(* IEC 61131-3 sources: plc-st-coding-agent/progress/evidence/f14_v5_public_pilot_20261112/jobs/custom_deepseek-v4pro, 22 files *)

(* ---- public-easy-01.candidate_01.st ---- *)
TYPE LineState :
(
    IDLE,
    CLEANING,
    FILLING,
    CAPPING,
    PACKING,
    COMPLETE
);
END_TYPE;

FUNCTION_BLOCK AutomatedFillingLine
VAR_INPUT
    bottleSensor : BOOL;
    cleaningConfirmButton : BOOL;
    fillingConfirmButton : BOOL;
    cappingConfirmButton : BOOL;
    packingConfirmButton : BOOL;
    finishedButton : BOOL;
END_VAR
VAR_OUTPUT
    Pump_Motor : BOOL;
    Filling_Valve : BOOL;
    Capping_Machine : BOOL;
    Packing_Machine : BOOL;
    Completion_Light : BOOL;
END_VAR
VAR
    cleaningEdge : R_TRIG;
    fillingEdge : R_TRIG;
    cappingEdge : R_TRIG;
    packingEdge : R_TRIG;
    finishedEdge : R_TRIG;
    currentState : LineState := LineState#IDLE;
END_VAR

(*
ENGINEERING_CONTRACT
- Pump_Motor: activated when bottleSensor TRUE and state=IDLE -> CLEANING; retained until cleaningConfirm edge (PUB003, PUB004).
  Deactivated on cleaningConfirm edge.
- Filling_Valve: activated on cleaningConfirm edge after cleaning; retained until fillingConfirm edge (PUB004, PUB005).
  Deactivated on fillingConfirm edge.
- Capping_Machine: activated on fillingConfirm edge; retained until cappingConfirm edge (PUB005, PUB006).
  Deactivated on cappingConfirm edge.
- Packing_Machine: activated on cappingConfirm edge; retained until packingConfirm edge (PUB006, PUB007).
  Deactivated on packingConfirm edge.
- Completion_Light: activated on packingConfirm edge; retained until finishedButton edge (PUB007, PUB008).
  Deactivated on finishedButton edge, which also resets state to IDLE for next bottle.
- Same-scan priority: state transitions evaluated sequentially in scan order; no simultaneous edge trigger priority specified.
- Units: BOOL levels only; no timing/modbus scaling.
*)

cleaningEdge(CLK := cleaningConfirmButton);
fillingEdge(CLK := fillingConfirmButton);
cappingEdge(CLK := cappingConfirmButton);
packingEdge(CLK := packingConfirmButton);
finishedEdge(CLK := finishedButton);

CASE currentState OF
    LineState#IDLE:
        Pump_Motor := FALSE;
        Filling_Valve := FALSE;
        Capping_Machine := FALSE;
        Packing_Machine := FALSE;
        Completion_Light := FALSE;

        IF bottleSensor THEN
            currentState := LineState#CLEANING;
            Pump_Motor := TRUE;
        END_IF;

    LineState#CLEANING:
        Pump_Motor := TRUE;
        Filling_Valve := FALSE;
        Capping_Machine := FALSE;
        Packing_Machine := FALSE;
        Completion_Light := FALSE;

        IF cleaningEdge.Q THEN
            Pump_Motor := FALSE;
            Filling_Valve := TRUE;
            currentState := LineState#FILLING;
        END_IF;

    LineState#FILLING:
        Pump_Motor := FALSE;
        Filling_Valve := TRUE;
        Capping_Machine := FALSE;
        Packing_Machine := FALSE;
        Completion_Light := FALSE;

        IF fillingEdge.Q THEN
            Filling_Valve := FALSE;
            Capping_Machine := TRUE;
            currentState := LineState#CAPPING;
        END_IF;

    LineState#CAPPING:
        Pump_Motor := FALSE;
        Filling_Valve := FALSE;
        Capping_Machine := TRUE;
        Packing_Machine := FALSE;
        Completion_Light := FALSE;

        IF cappingEdge.Q THEN
            Capping_Machine := FALSE;
            Packing_Machine := TRUE;
            currentState := LineState#PACKING;
        END_IF;

    LineState#PACKING:
        Pump_Motor := FALSE;
        Filling_Valve := FALSE;
        Capping_Machine := FALSE;
        Packing_Machine := TRUE;
        Completion_Light := FALSE;

        IF packingEdge.Q THEN
            Packing_Machine := FALSE;
            Completion_Light := TRUE;
            currentState := LineState#COMPLETE;
        END_IF;

    LineState#COMPLETE:
        Pump_Motor := FALSE;
        Filling_Valve := FALSE;
        Capping_Machine := FALSE;
        Packing_Machine := FALSE;
        Completion_Light := TRUE;

        IF finishedEdge.Q THEN
            Completion_Light := FALSE;
            currentState := LineState#IDLE;
        END_IF;
END_CASE;
END_FUNCTION_BLOCK

(* ---- public-easy-01.candidate_02.st ---- *)
(*
ENGINEERING_CONTRACT
- Pump_Motor: activated when bottleSensor TRUE and state=IDLE -> CLEANING; retained until cleaningConfirm edge (PUB003, PUB004).
  Deactivated on cleaningConfirm edge.
- Filling_Valve: activated on cleaningConfirm edge after cleaning; retained until fillingConfirm edge (PUB004, PUB005).
  Deactivated on fillingConfirm edge.
- Capping_Machine: activated on fillingConfirm edge; retained until cappingConfirm edge (PUB005, PUB006).
  Deactivated on cappingConfirm edge.
- Packing_Machine: activated on cappingConfirm edge; retained until packingConfirm edge (PUB006, PUB007).
  Deactivated on packingConfirm edge.
- Completion_Light: activated on packingConfirm edge; retained until finishedButton edge (PUB007, PUB008).
  Deactivated on finishedButton edge, which also resets state to IDLE for next bottle.
- Same-scan priority: no simultaneous edge trigger priority specified; transitions evaluated sequentially.
- Units: BOOL levels only.
*)

TYPE LineState :
(
    IDLE,
    CLEANING,
    FILLING,
    CAPPING,
    PACKING,
    COMPLETE
);
END_TYPE;

FUNCTION_BLOCK AutomatedFillingLine
VAR_INPUT
    bottleSensor : BOOL;
    cleaningConfirmButton : BOOL;
    fillingConfirmButton : BOOL;
    cappingConfirmButton : BOOL;
    packingConfirmButton : BOOL;
    finishedButton : BOOL;
END_VAR
VAR_OUTPUT
    Pump_Motor : BOOL;
    Filling_Valve : BOOL;
    Capping_Machine : BOOL;
    Packing_Machine : BOOL;
    Completion_Light : BOOL;
END_VAR
VAR
    cleaningEdge : R_TRIG;
    fillingEdge : R_TRIG;
    cappingEdge : R_TRIG;
    packingEdge : R_TRIG;
    finishedEdge : R_TRIG;
    currentState : LineState := IDLE;
END_VAR

cleaningEdge(CLK := cleaningConfirmButton);
fillingEdge(CLK := fillingConfirmButton);
cappingEdge(CLK := cappingConfirmButton);
packingEdge(CLK := packingConfirmButton);
finishedEdge(CLK := finishedButton);

CASE currentState OF
    IDLE:
        Pump_Motor := FALSE;
        Filling_Valve := FALSE;
        Capping_Machine := FALSE;
        Packing_Machine := FALSE;
        Completion_Light := FALSE;

        IF bottleSensor THEN
            currentState := CLEANING;
            Pump_Motor := TRUE;
        END_IF;

    CLEANING:
        Pump_Motor := TRUE;
        Filling_Valve := FALSE;
        Capping_Machine := FALSE;
        Packing_Machine := FALSE;
        Completion_Light := FALSE;

        IF cleaningEdge.Q THEN
            Pump_Motor := FALSE;
            Filling_Valve := TRUE;
            currentState := FILLING;
        END_IF;

    FILLING:
        Pump_Motor := FALSE;
        Filling_Valve := TRUE;
        Capping_Machine := FALSE;
        Packing_Machine := FALSE;
        Completion_Light := FALSE;

        IF fillingEdge.Q THEN
            Filling_Valve := FALSE;
            Capping_Machine := TRUE;
            currentState := CAPPING;
        END_IF;

    CAPPING:
        Pump_Motor := FALSE;
        Filling_Valve := FALSE;
        Capping_Machine := TRUE;
        Packing_Machine := FALSE;
        Completion_Light := FALSE;

        IF cappingEdge.Q THEN
            Capping_Machine := FALSE;
            Packing_Machine := TRUE;
            currentState := PACKING;
        END_IF;

    PACKING:
        Pump_Motor := FALSE;
        Filling_Valve := FALSE;
        Capping_Machine := FALSE;
        Packing_Machine := TRUE;
        Completion_Light := FALSE;

        IF packingEdge.Q THEN
            Packing_Machine := FALSE;
            Completion_Light := TRUE;
            currentState := COMPLETE;
        END_IF;

    COMPLETE:
        Pump_Motor := FALSE;
        Filling_Valve := FALSE;
        Capping_Machine := FALSE;
        Packing_Machine := FALSE;
        Completion_Light := TRUE;

        IF finishedEdge.Q THEN
            Completion_Light := FALSE;
            currentState := IDLE;
        END_IF;
END_CASE;

END_FUNCTION_BLOCK

(* ---- public-easy-01.raw_candidate_01.st ---- *)
TYPE LineState :
(
    IDLE,
    CLEANING,
    FILLING,
    CAPPING,
    PACKING,
    COMPLETE
);
END_TYPE

FUNCTION_BLOCK AutomatedFillingLine
VAR_INPUT
    bottleSensor : BOOL;
    cleaningConfirmButton : BOOL;
    fillingConfirmButton : BOOL;
    cappingConfirmButton : BOOL;
    packingConfirmButton : BOOL;
    finishedButton : BOOL;
END_VAR
VAR_OUTPUT
    Pump_Motor : BOOL;
    Filling_Valve : BOOL;
    Capping_Machine : BOOL;
    Packing_Machine : BOOL;
    Completion_Light : BOOL;
END_VAR
VAR
    cleaningEdge : R_TRIG;
    fillingEdge : R_TRIG;
    cappingEdge : R_TRIG;
    packingEdge : R_TRIG;
    finishedEdge : R_TRIG;
    currentState : LineState := LineState#IDLE;
END_VAR

(*
ENGINEERING_CONTRACT
- Pump_Motor: activated when bottleSensor TRUE and state=IDLE -> CLEANING; retained until cleaningConfirm edge (PUB003, PUB004).
  Deactivated on cleaningConfirm edge.
- Filling_Valve: activated on cleaningConfirm edge after cleaning; retained until fillingConfirm edge (PUB004, PUB005).
  Deactivated on fillingConfirm edge.
- Capping_Machine: activated on fillingConfirm edge; retained until cappingConfirm edge (PUB005, PUB006).
  Deactivated on cappingConfirm edge.
- Packing_Machine: activated on cappingConfirm edge; retained until packingConfirm edge (PUB006, PUB007).
  Deactivated on packingConfirm edge.
- Completion_Light: activated on packingConfirm edge; retained until finishedButton edge (PUB007, PUB008).
  Deactivated on finishedButton edge, which also resets state to IDLE for next bottle.
- Same-scan priority: state transitions evaluated sequentially in scan order; no simultaneous edge trigger priority specified.
- Units: BOOL levels only; no timing/modbus scaling.
*)

cleaningEdge(CLK := cleaningConfirmButton);
fillingEdge(CLK := fillingConfirmButton);
cappingEdge(CLK := cappingConfirmButton);
packingEdge(CLK := packingConfirmButton);
finishedEdge(CLK := finishedButton);

CASE currentState OF
    LineState#IDLE:
        Pump_Motor := FALSE;
        Filling_Valve := FALSE;
        Capping_Machine := FALSE;
        Packing_Machine := FALSE;
        Completion_Light := FALSE;

        IF bottleSensor THEN
            currentState := LineState#CLEANING;
            Pump_Motor := TRUE;
        END_IF;

    LineState#CLEANING:
        Pump_Motor := TRUE;
        Filling_Valve := FALSE;
        Capping_Machine := FALSE;
        Packing_Machine := FALSE;
        Completion_Light := FALSE;

        IF cleaningEdge.Q THEN
            Pump_Motor := FALSE;
            Filling_Valve := TRUE;
            currentState := LineState#FILLING;
        END_IF;

    LineState#FILLING:
        Pump_Motor := FALSE;
        Filling_Valve := TRUE;
        Capping_Machine := FALSE;
        Packing_Machine := FALSE;
        Completion_Light := FALSE;

        IF fillingEdge.Q THEN
            Filling_Valve := FALSE;
            Capping_Machine := TRUE;
            currentState := LineState#CAPPING;
        END_IF;

    LineState#CAPPING:
        Pump_Motor := FALSE;
        Filling_Valve := FALSE;
        Capping_Machine := TRUE;
        Packing_Machine := FALSE;
        Completion_Light := FALSE;

        IF cappingEdge.Q THEN
            Capping_Machine := FALSE;
            Packing_Machine := TRUE;
            currentState := LineState#PACKING;
        END_IF;

    LineState#PACKING:
        Pump_Motor := FALSE;
        Filling_Valve := FALSE;
        Capping_Machine := FALSE;
        Packing_Machine := TRUE;
        Completion_Light := FALSE;

        IF packingEdge.Q THEN
            Packing_Machine := FALSE;
            Completion_Light := TRUE;
            currentState := LineState#COMPLETE;
        END_IF;

    LineState#COMPLETE:
        Pump_Motor := FALSE;
        Filling_Valve := FALSE;
        Capping_Machine := FALSE;
        Packing_Machine := FALSE;
        Completion_Light := TRUE;

        IF finishedEdge.Q THEN
            Completion_Light := FALSE;
            currentState := LineState#IDLE;
        END_IF;
END_CASE;
END_FUNCTION_BLOCK

(* ---- public-easy-01.raw_candidate_02.st ---- *)
(*
ENGINEERING_CONTRACT
- Pump_Motor: activated when bottleSensor TRUE and state=IDLE -> CLEANING; retained until cleaningConfirm edge (PUB003, PUB004).
  Deactivated on cleaningConfirm edge.
- Filling_Valve: activated on cleaningConfirm edge after cleaning; retained until fillingConfirm edge (PUB004, PUB005).
  Deactivated on fillingConfirm edge.
- Capping_Machine: activated on fillingConfirm edge; retained until cappingConfirm edge (PUB005, PUB006).
  Deactivated on cappingConfirm edge.
- Packing_Machine: activated on cappingConfirm edge; retained until packingConfirm edge (PUB006, PUB007).
  Deactivated on packingConfirm edge.
- Completion_Light: activated on packingConfirm edge; retained until finishedButton edge (PUB007, PUB008).
  Deactivated on finishedButton edge, which also resets state to IDLE for next bottle.
- Same-scan priority: no simultaneous edge trigger priority specified; transitions evaluated sequentially.
- Units: BOOL levels only.
*)

TYPE LineState :
(
    IDLE,
    CLEANING,
    FILLING,
    CAPPING,
    PACKING,
    COMPLETE
);
END_TYPE

FUNCTION_BLOCK AutomatedFillingLine
VAR_INPUT
    bottleSensor : BOOL;
    cleaningConfirmButton : BOOL;
    fillingConfirmButton : BOOL;
    cappingConfirmButton : BOOL;
    packingConfirmButton : BOOL;
    finishedButton : BOOL;
END_VAR
VAR_OUTPUT
    Pump_Motor : BOOL;
    Filling_Valve : BOOL;
    Capping_Machine : BOOL;
    Packing_Machine : BOOL;
    Completion_Light : BOOL;
END_VAR
VAR
    cleaningEdge : R_TRIG;
    fillingEdge : R_TRIG;
    cappingEdge : R_TRIG;
    packingEdge : R_TRIG;
    finishedEdge : R_TRIG;
    currentState : LineState := IDLE;
END_VAR

cleaningEdge(CLK := cleaningConfirmButton);
fillingEdge(CLK := fillingConfirmButton);
cappingEdge(CLK := cappingConfirmButton);
packingEdge(CLK := packingConfirmButton);
finishedEdge(CLK := finishedButton);

CASE currentState OF
    IDLE:
        Pump_Motor := FALSE;
        Filling_Valve := FALSE;
        Capping_Machine := FALSE;
        Packing_Machine := FALSE;
        Completion_Light := FALSE;

        IF bottleSensor THEN
            currentState := CLEANING;
            Pump_Motor := TRUE;
        END_IF;

    CLEANING:
        Pump_Motor := TRUE;
        Filling_Valve := FALSE;
        Capping_Machine := FALSE;
        Packing_Machine := FALSE;
        Completion_Light := FALSE;

        IF cleaningEdge.Q THEN
            Pump_Motor := FALSE;
            Filling_Valve := TRUE;
            currentState := FILLING;
        END_IF;

    FILLING:
        Pump_Motor := FALSE;
        Filling_Valve := TRUE;
        Capping_Machine := FALSE;
        Packing_Machine := FALSE;
        Completion_Light := FALSE;

        IF fillingEdge.Q THEN
            Filling_Valve := FALSE;
            Capping_Machine := TRUE;
            currentState := CAPPING;
        END_IF;

    CAPPING:
        Pump_Motor := FALSE;
        Filling_Valve := FALSE;
        Capping_Machine := TRUE;
        Packing_Machine := FALSE;
        Completion_Light := FALSE;

        IF cappingEdge.Q THEN
            Capping_Machine := FALSE;
            Packing_Machine := TRUE;
            currentState := PACKING;
        END_IF;

    PACKING:
        Pump_Motor := FALSE;
        Filling_Valve := FALSE;
        Capping_Machine := FALSE;
        Packing_Machine := TRUE;
        Completion_Light := FALSE;

        IF packingEdge.Q THEN
            Packing_Machine := FALSE;
            Completion_Light := TRUE;
            currentState := COMPLETE;
        END_IF;

    COMPLETE:
        Pump_Motor := FALSE;
        Filling_Valve := FALSE;
        Capping_Machine := FALSE;
        Packing_Machine := FALSE;
        Completion_Light := TRUE;

        IF finishedEdge.Q THEN
            Completion_Light := FALSE;
            currentState := IDLE;
        END_IF;
END_CASE;

END_FUNCTION_BLOCK

(* ---- public-easy-04.candidate_01.st ---- *)
FUNCTION_BLOCK FB_JamPumpDebounceRuntime
VAR_INPUT
    VISCOSITY_OK : BOOL;
    PASTE_E_STOP_NC : BOOL;
    DebounceTime : TIME;
    CycleTime : TIME;
END_VAR
VAR_OUTPUT
    VFD_RUN : BOOL := FALSE;
    PUMP_MAINT_DUE : BOOL := FALSE;
    PUMP_RUNTIME_ACC : LTIME := LTIME#0s;
END_VAR
VAR
    DebounceTimer : TON;
    TonIn : BOOL;
    ViscosityValid : BOOL;
    AccRuntime : LTIME := LTIME#0s;
    MAINT_THRESHOLD : LTIME := LTIME#500h;
END_VAR

(*
ENGINEERING_CONTRACT:
- VFD_RUN activation: PASTE_E_STOP_NC AND ViscosityValid; no latch.
- ViscosityValid: TON Q; debounce reset when VISCOSITY_OK FALSE or E-STOP FALSE while incomplete (PUB002/PUB003).
- E-stop same-scan priority: VFD_RUN false if PASTE_E_STOP_NC false; incomplete timer cleared.
- PUMP_RUNTIME_ACC: retained while stopped; adds CycleTime only when VFD_RUN TRUE; init 0 (PUB004/PUB005).
- PUMP_MAINT_DUE: informational latch at >= LTIME#500h; does not affect VFD_RUN (PUB004/PUB005).
- Units: DebounceTime TIME ms, CycleTime TIME ms converted to LTIME ns; threshold 500h.
*)

TonIn := VISCOSITY_OK AND (PASTE_E_STOP_NC OR DebounceTimer.Q);
DebounceTimer(IN := TonIn, PT := DebounceTime);
ViscosityValid := DebounceTimer.Q;

VFD_RUN := PASTE_E_STOP_NC AND ViscosityValid;

IF VFD_RUN THEN
    AccRuntime := AccRuntime + TIME_TO_LTIME(CycleTime);
END_IF;

PUMP_RUNTIME_ACC := AccRuntime;
PUMP_MAINT_DUE := (AccRuntime >= MAINT_THRESHOLD);

END_FUNCTION_BLOCK

(* ---- public-easy-04.raw_candidate_01.st ---- *)
FUNCTION_BLOCK FB_JamPumpDebounceRuntime
VAR_INPUT
    VISCOSITY_OK : BOOL;
    PASTE_E_STOP_NC : BOOL;
    DebounceTime : TIME;
    CycleTime : TIME;
END_VAR
VAR_OUTPUT
    VFD_RUN : BOOL := FALSE;
    PUMP_MAINT_DUE : BOOL := FALSE;
    PUMP_RUNTIME_ACC : LTIME := LTIME#0s;
END_VAR
VAR
    DebounceTimer : TON;
    TonIn : BOOL;
    ViscosityValid : BOOL;
    AccRuntime : LTIME := LTIME#0s;
    MAINT_THRESHOLD : LTIME := LTIME#500h;
END_VAR

(*
ENGINEERING_CONTRACT:
- VFD_RUN activation: PASTE_E_STOP_NC AND ViscosityValid; no latch.
- ViscosityValid: TON Q; debounce reset when VISCOSITY_OK FALSE or E-STOP FALSE while incomplete (PUB002/PUB003).
- E-stop same-scan priority: VFD_RUN false if PASTE_E_STOP_NC false; incomplete timer cleared.
- PUMP_RUNTIME_ACC: retained while stopped; adds CycleTime only when VFD_RUN TRUE; init 0 (PUB004/PUB005).
- PUMP_MAINT_DUE: informational latch at >= LTIME#500h; does not affect VFD_RUN (PUB004/PUB005).
- Units: DebounceTime TIME ms, CycleTime TIME ms converted to LTIME ns; threshold 500h.
*)

TonIn := VISCOSITY_OK AND (PASTE_E_STOP_NC OR DebounceTimer.Q);
DebounceTimer(IN := TonIn, PT := DebounceTime);
ViscosityValid := DebounceTimer.Q;

VFD_RUN := PASTE_E_STOP_NC AND ViscosityValid;

IF VFD_RUN THEN
    AccRuntime := AccRuntime + TIME_TO_LTIME(CycleTime);
END_IF;

PUMP_RUNTIME_ACC := AccRuntime;
PUMP_MAINT_DUE := (AccRuntime >= MAINT_THRESHOLD);

END_FUNCTION_BLOCK

(* ---- public-hard-03.candidate_01.st ---- *)
TYPE ST_Recipe :
STRUCT
    recipeID : INT;
    ingredientType : INT;
    ingredientRatio : REAL;
    productionTemperature : REAL;
END_STRUCT
END_TYPE;

FUNCTION_BLOCK RecipeManagementSystem
VAR_INPUT
    addRecipe : BOOL;
    deleteRecipe : BOOL;
    modifyRecipe : BOOL;
    queryRecipe : BOOL;
    recipeIn : ST_Recipe;
END_VAR
VAR_OUTPUT
    recipeAdded : BOOL;
    recipeDeleted : BOOL;
    recipeModified : BOOL;
    recipeQueryResult : ST_Recipe;
    error : BOOL;
    status : WORD;
END_VAR
VAR_IN_OUT
    recipe : ARRAY[1..10] OF ST_Recipe;
END_VAR
VAR
    i : INT;
    foundIndex : INT;
    emptyIndex : INT;
    duplicate : BOOL;
END_VAR

(*
ENGINEERING_CONTRACT
- Commands are level-triggered and evaluated each scan. No edge detection.
- Priority when simultaneous: add > delete > modify > query (IF/ELSIF). Unspecified by task.
- Outputs default FALSE / 0 / zero recipe each scan. Success outputs pulse with command.
- error/status default no error (0); set to 16#8001..16#8005 on failure.
- recipeQueryResult zeroed unless query success; no separate query success output.
- recipe array is inout storage; add fills lowest recipeID=0 slot; delete sets recipeID=0 only; modify overwrites matched slot.
- recipeID=0 is reserved; query/delete/modify treat 0 as not found; add rejects 0 as duplicate/reserved (16#8002).
- Duplicate check ignores empty slots, but add 0 special-cased.
- PUB009-PUB012 define error codes and operations.
*)

(* Default outputs each scan *)
recipeAdded := FALSE;
recipeDeleted := FALSE;
recipeModified := FALSE;
error := FALSE;
status := WORD#16#0000;
recipeQueryResult.recipeID := 0;
recipeQueryResult.ingredientType := 0;
recipeQueryResult.ingredientRatio := 0.0;
recipeQueryResult.productionTemperature := 0.0;

(* Add recipe *)
IF addRecipe THEN
    duplicate := FALSE;
    emptyIndex := 0;

    (* recipeID=0 is reserved as empty slot; reject as duplicate *)
    IF recipeIn.recipeID = 0 THEN
        duplicate := TRUE;
    ELSE
        FOR i := 1 TO 10 DO
            IF (recipe[i].recipeID <> 0) AND (recipe[i].recipeID = recipeIn.recipeID) THEN
                duplicate := TRUE;
                EXIT;
            END_IF;
        END_FOR;
    END_IF;

    IF duplicate THEN
        error := TRUE;
        status := WORD#16#8002;
    ELSE
        (* Find smallest empty slot *)
        FOR i := 1 TO 10 DO
            IF recipe[i].recipeID = 0 THEN
                emptyIndex := i;
                EXIT;
            END_IF;
        END_FOR;

        IF emptyIndex = 0 THEN
            error := TRUE;
            status := WORD#16#8003;
        ELSE
            recipe[emptyIndex] := recipeIn;
            recipeAdded := TRUE;
        END_IF;
    END_IF;

(* Delete recipe *)
ELSIF deleteRecipe THEN
    foundIndex := 0;

    IF recipeIn.recipeID <> 0 THEN
        FOR i := 1 TO 10 DO
            IF (recipe[i].recipeID <> 0) AND (recipe[i].recipeID = recipeIn.recipeID) THEN
                foundIndex := i;
                EXIT;
            END_IF;
        END_FOR;
    END_IF;

    IF foundIndex = 0 THEN
        error := TRUE;
        status := WORD#16#8004;
    ELSE
        recipe[foundIndex].recipeID := 0;
        recipeDeleted := TRUE;
    END_IF;

(* Modify recipe *)
ELSIF modifyRecipe THEN
    foundIndex := 0;

    IF recipeIn.recipeID <> 0 THEN
        FOR i := 1 TO 10 DO
            IF (recipe[i].recipeID <> 0) AND (recipe[i].recipeID = recipeIn.recipeID) THEN
                foundIndex := i;
                EXIT;
            END_IF;
        END_FOR;
    END_IF;

    IF foundIndex = 0 THEN
        error := TRUE;
        status := WORD#16#8005;
    ELSE
        recipe[foundIndex] := recipeIn;
        recipeModified := TRUE;
    END_IF;

(* Query recipe *)
ELSIF queryRecipe THEN
    foundIndex := 0;

    IF recipeIn.recipeID <> 0 THEN
        FOR i := 1 TO 10 DO
            IF (recipe[i].recipeID <> 0) AND (recipe[i].recipeID = recipeIn.recipeID) THEN
                foundIndex := i;
                EXIT;
            END_IF;
        END_FOR;
    END_IF;

    IF foundIndex = 0 THEN
        error := TRUE;
        status := WORD#16#8001;
    ELSE
        recipeQueryResult := recipe[foundIndex];
    END_IF;
END_IF;

END_FUNCTION_BLOCK

(* ---- public-hard-03.candidate_02.st ---- *)
TYPE ST_Recipe :
STRUCT
    recipeID : INT;
    ingredientType : INT;
    ingredientRatio : REAL;
    productionTemperature : REAL;
END_STRUCT
END_TYPE;

FUNCTION_BLOCK RecipeManagementSystem
VAR_INPUT
    addRecipe : BOOL;
    deleteRecipe : BOOL;
    modifyRecipe : BOOL;
    queryRecipe : BOOL;
    recipeIn : ST_Recipe;
END_VAR
VAR_OUTPUT
    recipeAdded : BOOL;
    recipeDeleted : BOOL;
    recipeModified : BOOL;
    recipeQueryResult : ST_Recipe;
    error : BOOL;
    status : WORD;
END_VAR
VAR_IN_OUT
    recipe : ARRAY[1..10] OF ST_Recipe;
END_VAR
VAR
    trigAdd : R_TRIG;
    trigDelete : R_TRIG;
    trigModify : R_TRIG;
    trigQuery : R_TRIG;
    addPulse : BOOL;
    deletePulse : BOOL;
    modifyPulse : BOOL;
    queryPulse : BOOL;
    i : INT;
    foundIndex : INT;
    emptyIndex : INT;
    duplicate : BOOL;
END_VAR

(*
ENGINEERING_CONTRACT
- Commands are edge-triggered: only the rising edge of each request executes the operation once.
- Priority when simultaneous edges occur: add > delete > modify > query (IF/ELSIF chain). Unspecified by task.
- Default outputs: success flags FALSE, error FALSE, status 0, recipeQueryResult zeroed each scan.
- error/status remain FALSE/0 on success; set to 16#8001..16#8005 on respective failure.
- recipe array is persistent inout storage. Add fills the lowest recipeID=0 slot; delete sets recipeID=0 only; modify overwrites the matched slot with the full input recipe.
- recipeID=0 is reserved as empty; query/delete/modify treat 0 as “not found”; add rejects 0 with duplicate error 16#8002 (as it conflicts with empty slots).
- PUB009-PUB012 define error codes and operations.
*)

(* Rising-edge detection for all command inputs *)
trigAdd(CLK := addRecipe);
addPulse := trigAdd.Q;
trigDelete(CLK := deleteRecipe);
deletePulse := trigDelete.Q;
trigModify(CLK := modifyRecipe);
modifyPulse := trigModify.Q;
trigQuery(CLK := queryRecipe);
queryPulse := trigQuery.Q;

(* Default outputs each scan *)
recipeAdded := FALSE;
recipeDeleted := FALSE;
recipeModified := FALSE;
error := FALSE;
status := WORD#16#0000;
recipeQueryResult.recipeID := 0;
recipeQueryResult.ingredientType := 0;
recipeQueryResult.ingredientRatio := 0.0;
recipeQueryResult.productionTemperature := 0.0;

(* Add recipe *)
IF addPulse THEN
    duplicate := FALSE;
    emptyIndex := 0;

    (* recipeID=0 is reserved as empty slot; reject as duplicate *)
    IF recipeIn.recipeID = 0 THEN
        duplicate := TRUE;
    ELSE
        FOR i := 1 TO 10 DO
            IF (recipe[i].recipeID <> 0) AND (recipe[i].recipeID = recipeIn.recipeID) THEN
                duplicate := TRUE;
                EXIT;
            END_IF;
        END_FOR;
    END_IF;

    IF duplicate THEN
        error := TRUE;
        status := WORD#16#8002;
    ELSE
        (* Find smallest empty slot *)
        FOR i := 1 TO 10 DO
            IF recipe[i].recipeID = 0 THEN
                emptyIndex := i;
                EXIT;
            END_IF;
        END_FOR;

        IF emptyIndex = 0 THEN
            error := TRUE;
            status := WORD#16#8003;
        ELSE
            recipe[emptyIndex] := recipeIn;
            recipeAdded := TRUE;
        END_IF;
    END_IF;

(* Delete recipe *)
ELSIF deletePulse THEN
    foundIndex := 0;

    IF recipeIn.recipeID <> 0 THEN
        FOR i := 1 TO 10 DO
            IF (recipe[i].recipeID <> 0) AND (recipe[i].recipeID = recipeIn.recipeID) THEN
                foundIndex := i;
                EXIT;
            END_IF;
        END_FOR;
    END_IF;

    IF foundIndex = 0 THEN
        error := TRUE;
        status := WORD#16#8004;
    ELSE
        recipe[foundIndex].recipeID := 0;
        recipeDeleted := TRUE;
    END_IF;

(* Modify recipe *)
ELSIF modifyPulse THEN
    foundIndex := 0;

    IF recipeIn.recipeID <> 0 THEN
        FOR i := 1 TO 10 DO
            IF (recipe[i].recipeID <> 0) AND (recipe[i].recipeID = recipeIn.recipeID) THEN
                foundIndex := i;
                EXIT;
            END_IF;
        END_FOR;
    END_IF;

    IF foundIndex = 0 THEN
        error := TRUE;
        status := WORD#16#8005;
    ELSE
        recipe[foundIndex] := recipeIn;
        recipeModified := TRUE;
    END_IF;

(* Query recipe *)
ELSIF queryPulse THEN
    foundIndex := 0;

    IF recipeIn.recipeID <> 0 THEN
        FOR i := 1 TO 10 DO
            IF (recipe[i].recipeID <> 0) AND (recipe[i].recipeID = recipeIn.recipeID) THEN
                foundIndex := i;
                EXIT;
            END_IF;
        END_FOR;
    END_IF;

    IF foundIndex = 0 THEN
        error := TRUE;
        status := WORD#16#8001;
    ELSE
        recipeQueryResult := recipe[foundIndex];
    END_IF;
END_IF;

END_FUNCTION_BLOCK

(* ---- public-hard-03.raw_candidate_01.st ---- *)
TYPE ST_Recipe :
STRUCT
    recipeID : INT;
    ingredientType : INT;
    ingredientRatio : REAL;
    productionTemperature : REAL;
END_STRUCT
END_TYPE

FUNCTION_BLOCK RecipeManagementSystem
VAR_INPUT
    addRecipe : BOOL;
    deleteRecipe : BOOL;
    modifyRecipe : BOOL;
    queryRecipe : BOOL;
    recipeIn : ST_Recipe;
END_VAR
VAR_OUTPUT
    recipeAdded : BOOL;
    recipeDeleted : BOOL;
    recipeModified : BOOL;
    recipeQueryResult : ST_Recipe;
    error : BOOL;
    status : WORD;
END_VAR
VAR_IN_OUT
    recipe : ARRAY[1..10] OF ST_Recipe;
END_VAR
VAR
    i : INT;
    foundIndex : INT;
    emptyIndex : INT;
    duplicate : BOOL;
END_VAR

(*
ENGINEERING_CONTRACT
- Commands are level-triggered and evaluated each scan. No edge detection.
- Priority when simultaneous: add > delete > modify > query (IF/ELSIF). Unspecified by task.
- Outputs default FALSE / 0 / zero recipe each scan. Success outputs pulse with command.
- error/status default no error (0); set to 16#8001..16#8005 on failure.
- recipeQueryResult zeroed unless query success; no separate query success output.
- recipe array is inout storage; add fills lowest recipeID=0 slot; delete sets recipeID=0 only; modify overwrites matched slot.
- recipeID=0 is reserved; query/delete/modify treat 0 as not found; add rejects 0 as duplicate/reserved (16#8002).
- Duplicate check ignores empty slots, but add 0 special-cased.
- PUB009-PUB012 define error codes and operations.
*)

(* Default outputs each scan *)
recipeAdded := FALSE;
recipeDeleted := FALSE;
recipeModified := FALSE;
error := FALSE;
status := WORD#16#0000;
recipeQueryResult.recipeID := 0;
recipeQueryResult.ingredientType := 0;
recipeQueryResult.ingredientRatio := 0.0;
recipeQueryResult.productionTemperature := 0.0;

(* Add recipe *)
IF addRecipe THEN
    duplicate := FALSE;
    emptyIndex := 0;

    (* recipeID=0 is reserved as empty slot; reject as duplicate *)
    IF recipeIn.recipeID = 0 THEN
        duplicate := TRUE;
    ELSE
        FOR i := 1 TO 10 DO
            IF (recipe[i].recipeID <> 0) AND (recipe[i].recipeID = recipeIn.recipeID) THEN
                duplicate := TRUE;
                EXIT;
            END_IF;
        END_FOR;
    END_IF;

    IF duplicate THEN
        error := TRUE;
        status := WORD#16#8002;
    ELSE
        (* Find smallest empty slot *)
        FOR i := 1 TO 10 DO
            IF recipe[i].recipeID = 0 THEN
                emptyIndex := i;
                EXIT;
            END_IF;
        END_FOR;

        IF emptyIndex = 0 THEN
            error := TRUE;
            status := WORD#16#8003;
        ELSE
            recipe[emptyIndex] := recipeIn;
            recipeAdded := TRUE;
        END_IF;
    END_IF;

(* Delete recipe *)
ELSIF deleteRecipe THEN
    foundIndex := 0;

    IF recipeIn.recipeID <> 0 THEN
        FOR i := 1 TO 10 DO
            IF (recipe[i].recipeID <> 0) AND (recipe[i].recipeID = recipeIn.recipeID) THEN
                foundIndex := i;
                EXIT;
            END_IF;
        END_FOR;
    END_IF;

    IF foundIndex = 0 THEN
        error := TRUE;
        status := WORD#16#8004;
    ELSE
        recipe[foundIndex].recipeID := 0;
        recipeDeleted := TRUE;
    END_IF;

(* Modify recipe *)
ELSIF modifyRecipe THEN
    foundIndex := 0;

    IF recipeIn.recipeID <> 0 THEN
        FOR i := 1 TO 10 DO
            IF (recipe[i].recipeID <> 0) AND (recipe[i].recipeID = recipeIn.recipeID) THEN
                foundIndex := i;
                EXIT;
            END_IF;
        END_FOR;
    END_IF;

    IF foundIndex = 0 THEN
        error := TRUE;
        status := WORD#16#8005;
    ELSE
        recipe[foundIndex] := recipeIn;
        recipeModified := TRUE;
    END_IF;

(* Query recipe *)
ELSIF queryRecipe THEN
    foundIndex := 0;

    IF recipeIn.recipeID <> 0 THEN
        FOR i := 1 TO 10 DO
            IF (recipe[i].recipeID <> 0) AND (recipe[i].recipeID = recipeIn.recipeID) THEN
                foundIndex := i;
                EXIT;
            END_IF;
        END_FOR;
    END_IF;

    IF foundIndex = 0 THEN
        error := TRUE;
        status := WORD#16#8001;
    ELSE
        recipeQueryResult := recipe[foundIndex];
    END_IF;
END_IF;

END_FUNCTION_BLOCK

(* ---- public-hard-03.raw_candidate_02.st ---- *)
TYPE ST_Recipe :
STRUCT
    recipeID : INT;
    ingredientType : INT;
    ingredientRatio : REAL;
    productionTemperature : REAL;
END_STRUCT
END_TYPE;

FUNCTION_BLOCK RecipeManagementSystem
VAR_INPUT
    addRecipe : BOOL;
    deleteRecipe : BOOL;
    modifyRecipe : BOOL;
    queryRecipe : BOOL;
    recipeIn : ST_Recipe;
END_VAR
VAR_OUTPUT
    recipeAdded : BOOL;
    recipeDeleted : BOOL;
    recipeModified : BOOL;
    recipeQueryResult : ST_Recipe;
    error : BOOL;
    status : WORD;
END_VAR
VAR_IN_OUT
    recipe : ARRAY[1..10] OF ST_Recipe;
END_VAR
VAR
    trigAdd : R_TRIG;
    trigDelete : R_TRIG;
    trigModify : R_TRIG;
    trigQuery : R_TRIG;
    addPulse : BOOL;
    deletePulse : BOOL;
    modifyPulse : BOOL;
    queryPulse : BOOL;
    i : INT;
    foundIndex : INT;
    emptyIndex : INT;
    duplicate : BOOL;
END_VAR

(*
ENGINEERING_CONTRACT
- Commands are edge-triggered: only the rising edge of each request executes the operation once.
- Priority when simultaneous edges occur: add > delete > modify > query (IF/ELSIF chain). Unspecified by task.
- Default outputs: success flags FALSE, error FALSE, status 0, recipeQueryResult zeroed each scan.
- error/status remain FALSE/0 on success; set to 16#8001..16#8005 on respective failure.
- recipe array is persistent inout storage. Add fills the lowest recipeID=0 slot; delete sets recipeID=0 only; modify overwrites the matched slot with the full input recipe.
- recipeID=0 is reserved as empty; query/delete/modify treat 0 as “not found”; add rejects 0 with duplicate error 16#8002 (as it conflicts with empty slots).
- PUB009-PUB012 define error codes and operations.
*)

(* Rising-edge detection for all command inputs *)
trigAdd(CLK := addRecipe);
addPulse := trigAdd.Q;
trigDelete(CLK := deleteRecipe);
deletePulse := trigDelete.Q;
trigModify(CLK := modifyRecipe);
modifyPulse := trigModify.Q;
trigQuery(CLK := queryRecipe);
queryPulse := trigQuery.Q;

(* Default outputs each scan *)
recipeAdded := FALSE;
recipeDeleted := FALSE;
recipeModified := FALSE;
error := FALSE;
status := WORD#16#0000;
recipeQueryResult.recipeID := 0;
recipeQueryResult.ingredientType := 0;
recipeQueryResult.ingredientRatio := 0.0;
recipeQueryResult.productionTemperature := 0.0;

(* Add recipe *)
IF addPulse THEN
    duplicate := FALSE;
    emptyIndex := 0;

    (* recipeID=0 is reserved as empty slot; reject as duplicate *)
    IF recipeIn.recipeID = 0 THEN
        duplicate := TRUE;
    ELSE
        FOR i := 1 TO 10 DO
            IF (recipe[i].recipeID <> 0) AND (recipe[i].recipeID = recipeIn.recipeID) THEN
                duplicate := TRUE;
                EXIT;
            END_IF;
        END_FOR;
    END_IF;

    IF duplicate THEN
        error := TRUE;
        status := WORD#16#8002;
    ELSE
        (* Find smallest empty slot *)
        FOR i := 1 TO 10 DO
            IF recipe[i].recipeID = 0 THEN
                emptyIndex := i;
                EXIT;
            END_IF;
        END_FOR;

        IF emptyIndex = 0 THEN
            error := TRUE;
            status := WORD#16#8003;
        ELSE
            recipe[emptyIndex] := recipeIn;
            recipeAdded := TRUE;
        END_IF;
    END_IF;

(* Delete recipe *)
ELSIF deletePulse THEN
    foundIndex := 0;

    IF recipeIn.recipeID <> 0 THEN
        FOR i := 1 TO 10 DO
            IF (recipe[i].recipeID <> 0) AND (recipe[i].recipeID = recipeIn.recipeID) THEN
                foundIndex := i;
                EXIT;
            END_IF;
        END_FOR;
    END_IF;

    IF foundIndex = 0 THEN
        error := TRUE;
        status := WORD#16#8004;
    ELSE
        recipe[foundIndex].recipeID := 0;
        recipeDeleted := TRUE;
    END_IF;

(* Modify recipe *)
ELSIF modifyPulse THEN
    foundIndex := 0;

    IF recipeIn.recipeID <> 0 THEN
        FOR i := 1 TO 10 DO
            IF (recipe[i].recipeID <> 0) AND (recipe[i].recipeID = recipeIn.recipeID) THEN
                foundIndex := i;
                EXIT;
            END_IF;
        END_FOR;
    END_IF;

    IF foundIndex = 0 THEN
        error := TRUE;
        status := WORD#16#8005;
    ELSE
        recipe[foundIndex] := recipeIn;
        recipeModified := TRUE;
    END_IF;

(* Query recipe *)
ELSIF queryPulse THEN
    foundIndex := 0;

    IF recipeIn.recipeID <> 0 THEN
        FOR i := 1 TO 10 DO
            IF (recipe[i].recipeID <> 0) AND (recipe[i].recipeID = recipeIn.recipeID) THEN
                foundIndex := i;
                EXIT;
            END_IF;
        END_FOR;
    END_IF;

    IF foundIndex = 0 THEN
        error := TRUE;
        status := WORD#16#8001;
    ELSE
        recipeQueryResult := recipe[foundIndex];
    END_IF;
END_IF;

END_FUNCTION_BLOCK

(* ---- public-medium-03.candidate_01.st ---- *)
(*
ENGINEERING_CONTRACT
Activation: add sample each scan if cyclicExecution=TRUE; otherwise only on rising edge of trigger (PUB002, PUB003).
Reset priority: reset=TRUE clears history, average:=0, windowSizeReached:=FALSE before validation/add (PUB004).
Window validation: windowSize outside [1..100] sets error:=TRUE, status:=16#8200, windowSizeReached:=FALSE, and freezes calculation; average holds last valid output (PUB004/PUB007).
Same-scan: reset evaluated first, then window validation, then add; cyclicExecution suppresses trigger add but trigger edge is tracked for later cycles.
Retention: average/windowSizeReached hold between enabled samples; windowSizeReached becomes TRUE when stored count reaches windowSize.
Units/bounds: windowSize integer [1..100]; average LREAL; status WORD codes 16#0000 success, 16#8200 invalid window.
Unspecified: valid windowSize changes trim oldest stored samples to the new window without a separate reset.
*)
FUNCTION_BLOCK FB
VAR
    history : ARRAY[0..99] OF LREAL;
    count : INT := 0;
    oldestIdx : INT := 0;
    lastTrigger : BOOL := FALSE;
    i : INT;
    idx : INT;
    sum : LREAL;
    needAdd : BOOL;
    wsValid : BOOL;
END_VAR

IF reset THEN
    count := 0;
    oldestIdx := 0;
    average := 0.0;
    windowSizeReached := FALSE;
END_IF;

wsValid := (windowSize >= 1) AND (windowSize <= 100);

IF NOT wsValid THEN
    error := TRUE;
    status := 16#8200;
    windowSizeReached := FALSE;
ELSE
    error := FALSE;
    status := 16#0000;
    IF NOT reset THEN
        IF cyclicExecution THEN
            needAdd := TRUE;
        ELSE
            needAdd := trigger AND NOT lastTrigger;
        END_IF;
        IF needAdd THEN
            idx := (oldestIdx + count) MOD 100;
            history[idx] := value;
            IF count < 100 THEN
                count := count + 1;
            ELSE
                oldestIdx := (oldestIdx + 1) MOD 100;
            END_IF;
            WHILE count > windowSize DO
                oldestIdx := (oldestIdx + 1) MOD 100;
                count := count - 1;
            END_WHILE;
            IF count > 0 THEN
                sum := 0.0;
                FOR i := 0 TO count - 1 DO
                    idx := (oldestIdx + i) MOD 100;
                    sum := sum + history[idx];
                END_FOR;
                average := sum / INT_TO_LREAL(count);
            ELSE
                average := 0.0;
            END_IF;
            windowSizeReached := (count >= windowSize);
        END_IF;
    END_IF;
END_IF;

lastTrigger := trigger;
END_FUNCTION_BLOCK

(* ---- public-medium-03.candidate_02.st ---- *)
(*
ENGINEERING_CONTRACT
Activation: add sample each scan if cyclicExecution=TRUE; otherwise only on rising edge of trigger (PUB002, PUB003).
Reset priority: reset=TRUE clears history, average:=0, windowSizeReached:=FALSE before validation/add (PUB004).
Window validation: windowSize outside [1..100] sets error:=TRUE, status:=16#8200, windowSizeReached:=FALSE, and freezes calculation; average holds last valid output (PUB004/PUB007).
Same-scan: reset evaluated first, then window validation, then add; cyclicExecution suppresses trigger add but trigger edge is tracked for later cycles.
Retention: average/windowSizeReached hold between enabled samples; windowSizeReached becomes TRUE when stored count reaches windowSize.
Units/bounds: windowSize integer [1..100]; average LREAL; status WORD codes 16#0000 success, 16#8200 invalid window.
Unspecified: valid windowSize changes trim oldest stored samples to the new window without a separate reset.
*)
FUNCTION_BLOCK FB
VAR_INPUT
    cyclicExecution : BOOL;
    trigger : BOOL;
    value : LREAL;
    windowSize : INT;
    reset : BOOL;
END_VAR
VAR_OUTPUT
    average : LREAL;
    windowSizeReached : BOOL;
    error : BOOL;
    status : WORD;
END_VAR
VAR
    history : ARRAY[0..99] OF LREAL;
    count : INT := 0;
    oldestIdx : INT := 0;
    lastTrigger : BOOL := FALSE;
    i : INT;
    idx : INT;
    sum : LREAL;
    needAdd : BOOL;
    wsValid : BOOL;
END_VAR

IF reset THEN
    count := 0;
    oldestIdx := 0;
    average := 0.0;
    windowSizeReached := FALSE;
END_IF;

wsValid := (windowSize >= 1) AND (windowSize <= 100);

IF NOT wsValid THEN
    error := TRUE;
    status := 16#8200;
    windowSizeReached := FALSE;
ELSE
    error := FALSE;
    status := 16#0000;
    IF NOT reset THEN
        IF cyclicExecution THEN
            needAdd := TRUE;
        ELSE
            needAdd := trigger AND NOT lastTrigger;
        END_IF;
        IF needAdd THEN
            idx := (oldestIdx + count) MOD 100;
            history[idx] := value;
            IF count < 100 THEN
                count := count + 1;
            ELSE
                oldestIdx := (oldestIdx + 1) MOD 100;
            END_IF;
            WHILE count > windowSize DO
                oldestIdx := (oldestIdx + 1) MOD 100;
                count := count - 1;
            END_WHILE;
            IF count > 0 THEN
                sum := 0.0;
                FOR i := 0 TO count - 1 DO
                    idx := (oldestIdx + i) MOD 100;
                    sum := sum + history[idx];
                END_FOR;
                average := sum / INT_TO_LREAL(count);
            ELSE
                average := 0.0;
            END_IF;
            windowSizeReached := (count >= windowSize);
        END_IF;
    END_IF;
END_IF;

lastTrigger := trigger;
END_FUNCTION_BLOCK

(* ---- public-medium-03.raw_candidate_01.st ---- *)
(*
ENGINEERING_CONTRACT
Activation: add sample each scan if cyclicExecution=TRUE; otherwise only on rising edge of trigger (PUB002, PUB003).
Reset priority: reset=TRUE clears history, average:=0, windowSizeReached:=FALSE before validation/add (PUB004).
Window validation: windowSize outside [1..100] sets error:=TRUE, status:=16#8200, windowSizeReached:=FALSE, and freezes calculation; average holds last valid output (PUB004/PUB007).
Same-scan: reset evaluated first, then window validation, then add; cyclicExecution suppresses trigger add but trigger edge is tracked for later cycles.
Retention: average/windowSizeReached hold between enabled samples; windowSizeReached becomes TRUE when stored count reaches windowSize.
Units/bounds: windowSize integer [1..100]; average LREAL; status WORD codes 16#0000 success, 16#8200 invalid window.
Unspecified: valid windowSize changes trim oldest stored samples to the new window without a separate reset.
*)
FUNCTION_BLOCK FB
VAR
    history : ARRAY[0..99] OF LREAL;
    count : INT := 0;
    oldestIdx : INT := 0;
    lastTrigger : BOOL := FALSE;
    i : INT;
    idx : INT;
    sum : LREAL;
    needAdd : BOOL;
    wsValid : BOOL;
END_VAR

IF reset THEN
    count := 0;
    oldestIdx := 0;
    average := 0.0;
    windowSizeReached := FALSE;
END_IF;

wsValid := (windowSize >= 1) AND (windowSize <= 100);

IF NOT wsValid THEN
    error := TRUE;
    status := 16#8200;
    windowSizeReached := FALSE;
ELSE
    error := FALSE;
    status := 16#0000;
    IF NOT reset THEN
        IF cyclicExecution THEN
            needAdd := TRUE;
        ELSE
            needAdd := trigger AND NOT lastTrigger;
        END_IF;
        IF needAdd THEN
            idx := (oldestIdx + count) MOD 100;
            history[idx] := value;
            IF count < 100 THEN
                count := count + 1;
            ELSE
                oldestIdx := (oldestIdx + 1) MOD 100;
            END_IF;
            WHILE count > windowSize DO
                oldestIdx := (oldestIdx + 1) MOD 100;
                count := count - 1;
            END_WHILE;
            IF count > 0 THEN
                sum := 0.0;
                FOR i := 0 TO count - 1 DO
                    idx := (oldestIdx + i) MOD 100;
                    sum := sum + history[idx];
                END_FOR;
                average := sum / INT_TO_LREAL(count);
            ELSE
                average := 0.0;
            END_IF;
            windowSizeReached := (count >= windowSize);
        END_IF;
    END_IF;
END_IF;

lastTrigger := trigger;
END_FUNCTION_BLOCK

(* ---- public-medium-03.raw_candidate_02.st ---- *)
(*
ENGINEERING_CONTRACT
Activation: add sample each scan if cyclicExecution=TRUE; otherwise only on rising edge of trigger (PUB002, PUB003).
Reset priority: reset=TRUE clears history, average:=0, windowSizeReached:=FALSE before validation/add (PUB004).
Window validation: windowSize outside [1..100] sets error:=TRUE, status:=16#8200, windowSizeReached:=FALSE, and freezes calculation; average holds last valid output (PUB004/PUB007).
Same-scan: reset evaluated first, then window validation, then add; cyclicExecution suppresses trigger add but trigger edge is tracked for later cycles.
Retention: average/windowSizeReached hold between enabled samples; windowSizeReached becomes TRUE when stored count reaches windowSize.
Units/bounds: windowSize integer [1..100]; average LREAL; status WORD codes 16#0000 success, 16#8200 invalid window.
Unspecified: valid windowSize changes trim oldest stored samples to the new window without a separate reset.
*)
FUNCTION_BLOCK FB
VAR_INPUT
    cyclicExecution : BOOL;
    trigger : BOOL;
    value : LREAL;
    windowSize : INT;
    reset : BOOL;
END_VAR
VAR_OUTPUT
    average : LREAL;
    windowSizeReached : BOOL;
    error : BOOL;
    status : WORD;
END_VAR
VAR
    history : ARRAY[0..99] OF LREAL;
    count : INT := 0;
    oldestIdx : INT := 0;
    lastTrigger : BOOL := FALSE;
    i : INT;
    idx : INT;
    sum : LREAL;
    needAdd : BOOL;
    wsValid : BOOL;
END_VAR

IF reset THEN
    count := 0;
    oldestIdx := 0;
    average := 0.0;
    windowSizeReached := FALSE;
END_IF;

wsValid := (windowSize >= 1) AND (windowSize <= 100);

IF NOT wsValid THEN
    error := TRUE;
    status := 16#8200;
    windowSizeReached := FALSE;
ELSE
    error := FALSE;
    status := 16#0000;
    IF NOT reset THEN
        IF cyclicExecution THEN
            needAdd := TRUE;
        ELSE
            needAdd := trigger AND NOT lastTrigger;
        END_IF;
        IF needAdd THEN
            idx := (oldestIdx + count) MOD 100;
            history[idx] := value;
            IF count < 100 THEN
                count := count + 1;
            ELSE
                oldestIdx := (oldestIdx + 1) MOD 100;
            END_IF;
            WHILE count > windowSize DO
                oldestIdx := (oldestIdx + 1) MOD 100;
                count := count - 1;
            END_WHILE;
            IF count > 0 THEN
                sum := 0.0;
                FOR i := 0 TO count - 1 DO
                    idx := (oldestIdx + i) MOD 100;
                    sum := sum + history[idx];
                END_FOR;
                average := sum / INT_TO_LREAL(count);
            ELSE
                average := 0.0;
            END_IF;
            windowSizeReached := (count >= windowSize);
        END_IF;
    END_IF;
END_IF;

lastTrigger := trigger;
END_FUNCTION_BLOCK

(* ---- public-medium-04.candidate_01.st ---- *)
FUNCTION_BLOCK FB_TemperatureControl
(* ENGINEERING_CONTRACT
   - CurrentTemperature: raw TemperatureSensorInput assigned every scan; no unit conversion; no retention.
   - SetTempDisplay: echoes SetTemperature every scan; no units/bounds applied.
   - HeaterStatus: equals HeaterOutput after all gating; no independent latch.
   - OverheatProtection: latched TRUE when continuous heater on-time exceeds 5 s (PUB006);
     cleared only after 3 s cooldown timer expires (PUB006); retains state across scans.
   - HeaterOutput: TRUE when sensor valid, not overheat-latched, and TemperatureSensorInput < SetTemperature (PUB003);
     FALSE when actual > set, equal, sensor fault, or overheat latched (PUB004/PUB005/PUB008).
   - Sensor fault: TemperatureSensorInput < 0.0 OR > 100.0 disables heating; non-latching (PUB008).
   - Boundary equality: heater off (unspecified by PUB003/PUB004; implemented consistently).
*)
VAR_INPUT
    TemperatureSensorInput : REAL;
    SetTemperature : REAL;
END_VAR
VAR_OUTPUT
    CurrentTemperature : REAL;
    SetTempDisplay : REAL;
    HeaterStatus : BOOL;
    OverheatProtection : BOOL;
    HeaterOutput : BOOL;
END_VAR
VAR
    sensorFault : BOOL;
    heaterCmd : BOOL;
    overheatLatched : BOOL;
    heatTimer : TON;
    coolTimer : TON;
END_VAR

CurrentTemperature := TemperatureSensorInput;
SetTempDisplay := SetTemperature;

sensorFault := (TemperatureSensorInput < 0.0) OR (TemperatureSensorInput > 100.0);

heaterCmd := FALSE;
IF NOT sensorFault THEN
    IF TemperatureSensorInput < SetTemperature THEN
        heaterCmd := TRUE;
    ELSIF TemperatureSensorInput > SetTemperature THEN
        heaterCmd := FALSE;
    ELSE
        heaterCmd := FALSE; (* equality -> OFF *)
    END_IF;
END_IF;

heatTimer(IN := heaterCmd AND NOT overheatLatched, PT := T#5S);
IF heatTimer.Q THEN
    overheatLatched := TRUE;
END_IF;

coolTimer(IN := overheatLatched, PT := T#3S);
IF coolTimer.Q THEN
    overheatLatched := FALSE;
END_IF;

OverheatProtection := overheatLatched;

IF sensorFault OR overheatLatched THEN
    HeaterOutput := FALSE;
ELSE
    HeaterOutput := heaterCmd;
END_IF;

HeaterStatus := HeaterOutput;

END_FUNCTION_BLOCK

(* ---- public-medium-04.candidate_02.st ---- *)
FUNCTION_BLOCK FB_TemperatureControl
(* ENGINEERING_CONTRACT
   - CurrentTemperature: raw TemperatureSensorInput assigned every scan; no unit conversion; no retention.
   - SetTempDisplay: echoes SetTemperature every scan; no units/bounds applied.
   - HeaterStatus: equals HeaterOutput after all gating; no independent latch.
   - OverheatProtection: latched TRUE when continuous heater on-time exceeds 5 s (PUB006);
     cleared only after 3 s cooldown timer expires (PUB006); retains state across scans.
   - HeaterOutput: TRUE when sensor valid, not overheat-latched, and TemperatureSensorInput < SetTemperature (PUB003);
     FALSE when actual > set, equal, sensor fault, or overheat latched (PUB004/PUB005/PUB008).
   - Sensor fault: TemperatureSensorInput < 0.0 OR > 100.0 disables heating; non-latching (PUB008).
   - Boundary equality: heater off (unspecified by PUB003/PUB004; implemented consistently).
   - Overheat trigger uses strict > 5s via heatTimer.ET > T#5S (PUB006: "more than a certain period").
*)
VAR_INPUT
    TemperatureSensorInput : REAL;
    SetTemperature : REAL;
END_VAR
VAR_OUTPUT
    CurrentTemperature : REAL;
    SetTempDisplay : REAL;
    HeaterStatus : BOOL;
    OverheatProtection : BOOL;
    HeaterOutput : BOOL;
END_VAR
VAR
    sensorFault : BOOL;
    heaterCmd : BOOL;
    overheatLatched : BOOL;
    heatTimer : TON;
    coolTimer : TON;
END_VAR

CurrentTemperature := TemperatureSensorInput;
SetTempDisplay := SetTemperature;

sensorFault := (TemperatureSensorInput < 0.0) OR (TemperatureSensorInput > 100.0);

heaterCmd := FALSE;
IF NOT sensorFault THEN
    IF TemperatureSensorInput < SetTemperature THEN
        heaterCmd := TRUE;
    ELSIF TemperatureSensorInput > SetTemperature THEN
        heaterCmd := FALSE;
    ELSE
        heaterCmd := FALSE; (* equality -> OFF *)
    END_IF;
END_IF;

(* Heat timer with PT > 5s so we can check strictly greater than 5 seconds *)
heatTimer(IN := heaterCmd AND NOT overheatLatched, PT := T#10S);
IF heatTimer.ET > T#5S THEN
    overheatLatched := TRUE;
END_IF;

(* Cooldown timer: 3 seconds before lifting protection *)
coolTimer(IN := overheatLatched, PT := T#3S);
IF coolTimer.Q THEN
    overheatLatched := FALSE;
END_IF;

OverheatProtection := overheatLatched;

IF sensorFault OR overheatLatched THEN
    HeaterOutput := FALSE;
ELSE
    HeaterOutput := heaterCmd;
END_IF;

HeaterStatus := HeaterOutput;

END_FUNCTION_BLOCK

(* ---- public-medium-04.raw_candidate_01.st ---- *)
FUNCTION_BLOCK FB_TemperatureControl
(* ENGINEERING_CONTRACT
   - CurrentTemperature: raw TemperatureSensorInput assigned every scan; no unit conversion; no retention.
   - SetTempDisplay: echoes SetTemperature every scan; no units/bounds applied.
   - HeaterStatus: equals HeaterOutput after all gating; no independent latch.
   - OverheatProtection: latched TRUE when continuous heater on-time exceeds 5 s (PUB006);
     cleared only after 3 s cooldown timer expires (PUB006); retains state across scans.
   - HeaterOutput: TRUE when sensor valid, not overheat-latched, and TemperatureSensorInput < SetTemperature (PUB003);
     FALSE when actual > set, equal, sensor fault, or overheat latched (PUB004/PUB005/PUB008).
   - Sensor fault: TemperatureSensorInput < 0.0 OR > 100.0 disables heating; non-latching (PUB008).
   - Boundary equality: heater off (unspecified by PUB003/PUB004; implemented consistently).
*)
VAR_INPUT
    TemperatureSensorInput : REAL;
    SetTemperature : REAL;
END_VAR
VAR_OUTPUT
    CurrentTemperature : REAL;
    SetTempDisplay : REAL;
    HeaterStatus : BOOL;
    OverheatProtection : BOOL;
    HeaterOutput : BOOL;
END_VAR
VAR
    sensorFault : BOOL;
    heaterCmd : BOOL;
    overheatLatched : BOOL;
    heatTimer : TON;
    coolTimer : TON;
END_VAR

CurrentTemperature := TemperatureSensorInput;
SetTempDisplay := SetTemperature;

sensorFault := (TemperatureSensorInput < 0.0) OR (TemperatureSensorInput > 100.0);

heaterCmd := FALSE;
IF NOT sensorFault THEN
    IF TemperatureSensorInput < SetTemperature THEN
        heaterCmd := TRUE;
    ELSIF TemperatureSensorInput > SetTemperature THEN
        heaterCmd := FALSE;
    ELSE
        heaterCmd := FALSE; (* equality -> OFF *)
    END_IF
END_IF

heatTimer(IN := heaterCmd AND NOT overheatLatched, PT := T#5S);
IF heatTimer.Q THEN
    overheatLatched := TRUE;
END_IF

coolTimer(IN := overheatLatched, PT := T#3S);
IF coolTimer.Q THEN
    overheatLatched := FALSE;
END_IF

OverheatProtection := overheatLatched;

IF sensorFault OR overheatLatched THEN
    HeaterOutput := FALSE;
ELSE
    HeaterOutput := heaterCmd;
END_IF

HeaterStatus := HeaterOutput;

END_FUNCTION_BLOCK

(* ---- public-medium-04.raw_candidate_02.st ---- *)
FUNCTION_BLOCK FB_TemperatureControl
(* ENGINEERING_CONTRACT
   - CurrentTemperature: raw TemperatureSensorInput assigned every scan; no unit conversion; no retention.
   - SetTempDisplay: echoes SetTemperature every scan; no units/bounds applied.
   - HeaterStatus: equals HeaterOutput after all gating; no independent latch.
   - OverheatProtection: latched TRUE when continuous heater on-time exceeds 5 s (PUB006);
     cleared only after 3 s cooldown timer expires (PUB006); retains state across scans.
   - HeaterOutput: TRUE when sensor valid, not overheat-latched, and TemperatureSensorInput < SetTemperature (PUB003);
     FALSE when actual > set, equal, sensor fault, or overheat latched (PUB004/PUB005/PUB008).
   - Sensor fault: TemperatureSensorInput < 0.0 OR > 100.0 disables heating; non-latching (PUB008).
   - Boundary equality: heater off (unspecified by PUB003/PUB004; implemented consistently).
   - Overheat trigger uses strict > 5s via heatTimer.ET > T#5S (PUB006: "more than a certain period").
*)
VAR_INPUT
    TemperatureSensorInput : REAL;
    SetTemperature : REAL;
END_VAR
VAR_OUTPUT
    CurrentTemperature : REAL;
    SetTempDisplay : REAL;
    HeaterStatus : BOOL;
    OverheatProtection : BOOL;
    HeaterOutput : BOOL;
END_VAR
VAR
    sensorFault : BOOL;
    heaterCmd : BOOL;
    overheatLatched : BOOL;
    heatTimer : TON;
    coolTimer : TON;
END_VAR

CurrentTemperature := TemperatureSensorInput;
SetTempDisplay := SetTemperature;

sensorFault := (TemperatureSensorInput < 0.0) OR (TemperatureSensorInput > 100.0);

heaterCmd := FALSE;
IF NOT sensorFault THEN
    IF TemperatureSensorInput < SetTemperature THEN
        heaterCmd := TRUE;
    ELSIF TemperatureSensorInput > SetTemperature THEN
        heaterCmd := FALSE;
    ELSE
        heaterCmd := FALSE; (* equality -> OFF *)
    END_IF;
END_IF;

(* Heat timer with PT > 5s so we can check strictly greater than 5 seconds *)
heatTimer(IN := heaterCmd AND NOT overheatLatched, PT := T#10S);
IF heatTimer.ET > T#5S THEN
    overheatLatched := TRUE;
END_IF;

(* Cooldown timer: 3 seconds before lifting protection *)
coolTimer(IN := overheatLatched, PT := T#3S);
IF coolTimer.Q THEN
    overheatLatched := FALSE;
END_IF;

OverheatProtection := overheatLatched;

IF sensorFault OR overheatLatched THEN
    HeaterOutput := FALSE;
ELSE
    HeaterOutput := heaterCmd;
END_IF;

HeaterStatus := HeaterOutput;

END_FUNCTION_BLOCK

(* ---- public-medium-08.candidate_01.st ---- *)
FUNCTION_BLOCK FB_IPv4Parser
VAR_INPUT
    ipText : STRING(254);
END_VAR
VAR_OUTPUT
    ipValue : UDINT;
END_VAR
VAR
    i : INT;
    len : INT;
    digit : INT;
    segVal : UDINT;
    segCount : INT;
    segHasDigit : BOOL;
END_VAR

(*
ENGINEERING_CONTRACT
- ipValue: activated on valid 4-segment parse (PUB001/PUB003); recomputed every scan, no retention.
- ipValue reset/deactivated: malformed/non-digit/incorrect segment count/out-of-range -> 0 (PUB004); first failing check returns immediately.
- Same-scan priority: pure combinational; default 0, valid path overwrites with assembled value; any invalid path assigns 0 then RETURN.
- Units/boundaries: UDINT output 0..4294967295; each segment 0..255; first segment MSB, fourth LSB (PUB003).
- segCount: local state; reset to 0 each call; increments on completed segment; success requires exactly 4 (PUB002).
- segHasDigit: local state; reset FALSE each call and after each period; must be TRUE before every segment boundary (PUB002).
- Unspecified: leading zeros are accepted as ordinary decimal digits; no leading-zero rejection stated.
*)

ipValue := 0;
segVal := 0;
segCount := 0;
segHasDigit := FALSE;
len := LEN(ipText);

FOR i := 1 TO len DO
    digit := BYTE_TO_INT(ipText[i]);

    IF (digit >= 48) AND (digit <= 57) THEN
        segVal := segVal * UDINT#10 + INT_TO_UDINT(digit - INT#48);
        IF segVal > 255 THEN
            ipValue := 0;
            RETURN;
        END_IF;
        segHasDigit := TRUE;

    ELSIF digit = 46 THEN
        IF NOT segHasDigit THEN
            ipValue := 0;
            RETURN;
        END_IF;

        ipValue := SHL(ipValue, UINT#8);
        ipValue := ipValue OR segVal;

        segCount := segCount + 1;
        IF segCount > 3 THEN
            ipValue := 0;
            RETURN;
        END_IF;

        segVal := 0;
        segHasDigit := FALSE;

    ELSE
        ipValue := 0;
        RETURN;
    END_IF;
END_FOR;

IF NOT segHasDigit THEN
    ipValue := 0;
    RETURN;
END_IF;

ipValue := SHL(ipValue, UINT#8);
ipValue := ipValue OR segVal;
segCount := segCount + 1;

IF segCount <> 4 THEN
    ipValue := 0;
    RETURN;
END_IF;

END_FUNCTION_BLOCK

(* ---- public-medium-08.candidate_02.st ---- *)
FUNCTION_BLOCK FB_IPv4Parser
VAR_INPUT
    ipText : STRING(254);
END_VAR
VAR_OUTPUT
    ipValue : UDINT;
END_VAR
VAR
    i : INT;
    digit : INT;
    segVal : UDINT;
    segCount : INT;
    segHasDigit : BOOL;
END_VAR

(*
ENGINEERING_CONTRACT
- ipValue: active only on valid 4-segment IPv4; recomputed every scan, no retention (PUB001/PUB003).
- ipValue reset: any malformed / nondigit / wrong segment count / out-of-range segment forces 0 immediately (PUB004).
- Same-scan priority: combinational; initializes ipValue=0, valid path overwrites; invalid path sets 0 then RETURN.
- Units/boundaries: UDINT output 0..4294967295; each segment 0..255; first segment MSB, fourth LSB (PUB003).
- segCount: local; reset to 0 each call; increments after each period and after last segment; success requires exactly 4 (PUB002).
- segHasDigit: local; reset FALSE each call and after each period; must be TRUE before every segment boundary and at end (PUB002).
- Unspecified: leading zeros accepted as plain decimal digits; no leading‑zero rejection stated.
*)

ipValue := 0;
segVal := 0;
segCount := 0;
segHasDigit := FALSE;
i := 1;

WHILE (i <= 254) AND (BYTE_TO_INT(ipText[i]) <> 0) DO
    digit := BYTE_TO_INT(ipText[i]);

    IF (digit >= 48) AND (digit <= 57) THEN
        segVal := segVal * UDINT#10 + INT_TO_UDINT(digit - INT#48);
        IF segVal > 255 THEN
            ipValue := 0;
            RETURN;
        END_IF;
        segHasDigit := TRUE;

    ELSIF digit = 46 THEN  (* '.' *)
        IF NOT segHasDigit THEN
            ipValue := 0;
            RETURN;
        END_IF;

        ipValue := SHL(ipValue, UINT#8);
        ipValue := ipValue OR segVal;

        segCount := segCount + 1;
        IF segCount > 3 THEN
            ipValue := 0;
            RETURN;
        END_IF;

        segVal := 0;
        segHasDigit := FALSE;

    ELSE
        ipValue := 0;
        RETURN;
    END_IF;

    i := i + 1;
END_WHILE;

IF NOT segHasDigit THEN
    ipValue := 0;
    RETURN;
END_IF;

ipValue := SHL(ipValue, UINT#8);
ipValue := ipValue OR segVal;
segCount := segCount + 1;

IF segCount <> 4 THEN
    ipValue := 0;
    RETURN;
END_IF;

END_FUNCTION_BLOCK

(* ---- public-medium-08.raw_candidate_01.st ---- *)
FUNCTION_BLOCK FB_IPv4Parser
VAR_INPUT
    ipText : STRING(254);
END_VAR
VAR_OUTPUT
    ipValue : UDINT;
END_VAR
VAR
    i : INT;
    len : INT;
    digit : INT;
    segVal : UDINT;
    segCount : INT;
    segHasDigit : BOOL;
END_VAR

(*
ENGINEERING_CONTRACT
- ipValue: activated on valid 4-segment parse (PUB001/PUB003); recomputed every scan, no retention.
- ipValue reset/deactivated: malformed/non-digit/incorrect segment count/out-of-range -> 0 (PUB004); first failing check returns immediately.
- Same-scan priority: pure combinational; default 0, valid path overwrites with assembled value; any invalid path assigns 0 then RETURN.
- Units/boundaries: UDINT output 0..4294967295; each segment 0..255; first segment MSB, fourth LSB (PUB003).
- segCount: local state; reset to 0 each call; increments on completed segment; success requires exactly 4 (PUB002).
- segHasDigit: local state; reset FALSE each call and after each period; must be TRUE before every segment boundary (PUB002).
- Unspecified: leading zeros are accepted as ordinary decimal digits; no leading-zero rejection stated.
*)

ipValue := 0;
segVal := 0;
segCount := 0;
segHasDigit := FALSE;
len := LEN(ipText);

FOR i := 1 TO len DO
    digit := BYTE_TO_INT(ipText[i]);

    IF (digit >= 48) AND (digit <= 57) THEN
        segVal := segVal * UDINT#10 + INT_TO_UDINT(digit - INT#48);
        IF segVal > 255 THEN
            ipValue := 0;
            RETURN;
        END_IF;
        segHasDigit := TRUE;

    ELSIF digit = 46 THEN
        IF NOT segHasDigit THEN
            ipValue := 0;
            RETURN;
        END_IF;

        ipValue := SHL(ipValue, UINT#8);
        ipValue := ipValue OR segVal;

        segCount := segCount + 1;
        IF segCount > 3 THEN
            ipValue := 0;
            RETURN;
        END_IF;

        segVal := 0;
        segHasDigit := FALSE;

    ELSE
        ipValue := 0;
        RETURN;
    END_IF;
END_FOR;

IF NOT segHasDigit THEN
    ipValue := 0;
    RETURN;
END_IF;

ipValue := SHL(ipValue, UINT#8);
ipValue := ipValue OR segVal;
segCount := segCount + 1;

IF segCount <> 4 THEN
    ipValue := 0;
    RETURN;
END_IF;

END_FUNCTION_BLOCK

(* ---- public-medium-08.raw_candidate_02.st ---- *)
FUNCTION_BLOCK FB_IPv4Parser
VAR_INPUT
    ipText : STRING(254);
END_VAR
VAR_OUTPUT
    ipValue : UDINT;
END_VAR
VAR
    i : INT;
    digit : INT;
    segVal : UDINT;
    segCount : INT;
    segHasDigit : BOOL;
END_VAR

(*
ENGINEERING_CONTRACT
- ipValue: active only on valid 4-segment IPv4; recomputed every scan, no retention (PUB001/PUB003).
- ipValue reset: any malformed / nondigit / wrong segment count / out-of-range segment forces 0 immediately (PUB004).
- Same-scan priority: combinational; initializes ipValue=0, valid path overwrites; invalid path sets 0 then RETURN.
- Units/boundaries: UDINT output 0..4294967295; each segment 0..255; first segment MSB, fourth LSB (PUB003).
- segCount: local; reset to 0 each call; increments after each period and after last segment; success requires exactly 4 (PUB002).
- segHasDigit: local; reset FALSE each call and after each period; must be TRUE before every segment boundary and at end (PUB002).
- Unspecified: leading zeros accepted as plain decimal digits; no leading‑zero rejection stated.
*)

ipValue := 0;
segVal := 0;
segCount := 0;
segHasDigit := FALSE;
i := 1;

WHILE (i <= 254) AND (BYTE_TO_INT(ipText[i]) <> 0) DO
    digit := BYTE_TO_INT(ipText[i]);

    IF (digit >= 48) AND (digit <= 57) THEN
        segVal := segVal * UDINT#10 + INT_TO_UDINT(digit - INT#48);
        IF segVal > 255 THEN
            ipValue := 0;
            RETURN;
        END_IF;
        segHasDigit := TRUE;

    ELSIF digit = 46 THEN  (* '.' *)
        IF NOT segHasDigit THEN
            ipValue := 0;
            RETURN;
        END_IF;

        ipValue := SHL(ipValue, UINT#8);
        ipValue := ipValue OR segVal;

        segCount := segCount + 1;
        IF segCount > 3 THEN
            ipValue := 0;
            RETURN;
        END_IF;

        segVal := 0;
        segHasDigit := FALSE;

    ELSE
        ipValue := 0;
        RETURN;
    END_IF;

    i := i + 1;
END_WHILE;

IF NOT segHasDigit THEN
    ipValue := 0;
    RETURN;
END_IF;

ipValue := SHL(ipValue, UINT#8);
ipValue := ipValue OR segVal;
segCount := segCount + 1;

IF segCount <> 4 THEN
    ipValue := 0;
    RETURN;
END_IF;

END_FUNCTION_BLOCK
